Fanuc KAREL source: KT00906.KL

PROGRAM KT00906
%NOLOCKGROUP
%ENVIRONMENT VECTR
VAR
  P1: JOINTPOS
  P2: JOINTPOS
  OUT: VECTOR
BEGIN
  OUT = APPROACH(P1)
END KT00906
